// FB_TaktGenerator: 脉冲发生器
// 描述: 生成固定频率的方波脉冲信号 (50%占空比)

FUNCTION_BLOCK FB_TaktGenerator
VAR_INPUT
    Enable : BOOL;   // 使能信号 (TRUE=启用脉冲输出)
END_VAR
VAR_OUTPUT
    Takt_10Hz    : BOOL;  // 10Hz脉冲输出 (周期100ms)
    Takt_5Hz     : BOOL;  // 5Hz脉冲输出 (周期200ms)
    Takt_2_5Hz   : BOOL;  // 2.5Hz脉冲输出 (周期400ms)
    Takt_2Hz     : BOOL;  // 2Hz脉冲输出 (周期500ms)
    Takt_1_25Hz  : BOOL;  // 1.25Hz脉冲输出 (周期800ms)
    Takt_1Hz     : BOOL;  // 1Hz脉冲输出 (周期1s)
    Takt_0_625Hz : BOOL;  // 0.625Hz脉冲输出 (周期1.6s)
    Takt_0_5Hz   : BOOL;  // 0.5Hz脉冲输出 (周期2s)
    Takt_0_25Hz  : BOOL;  // 0.25Hz脉冲输出 (周期4s)
    Takt_0_2Hz   : BOOL;  // 0.2Hz脉冲输出 (周期5s)
END_VAR
VAR
    Cnt_10Hz     : DINT := 0;
    Cnt_5Hz      : DINT := 0;
    Cnt_2_5Hz    : DINT := 0;
    Cnt_2Hz      : DINT := 0;
    Cnt_1_25Hz   : DINT := 0;
    Cnt_1Hz      : DINT := 0;
    Cnt_0_625Hz  : DINT := 0;
    Cnt_0_5Hz    : DINT := 0;
    Cnt_0_25Hz   : DINT := 0;
    Cnt_0_2Hz    : DINT := 0;
END_VAR

BEGIN
    IF #Enable THEN
        // 10Hz: 周期100ms (假设10ms/扫描周期, 半周期=5)
        #Cnt_10Hz := #Cnt_10Hz + 1;
        IF #Cnt_10Hz >= 5 THEN
            #Takt_10Hz := NOT #Takt_10Hz;
            #Cnt_10Hz := 0;
        END_IF;

        // 5Hz: 周期200ms (半周期=10)
        #Cnt_5Hz := #Cnt_5Hz + 1;
        IF #Cnt_5Hz >= 10 THEN
            #Takt_5Hz := NOT #Takt_5Hz;
            #Cnt_5Hz := 0;
        END_IF;

        // 2.5Hz: 周期400ms (半周期=20)
        #Cnt_2_5Hz := #Cnt_2_5Hz + 1;
        IF #Cnt_2_5Hz >= 20 THEN
            #Takt_2_5Hz := NOT #Takt_2_5Hz;
            #Cnt_2_5Hz := 0;
        END_IF;

        // 2Hz: 周期500ms (半周期=25)
        #Cnt_2Hz := #Cnt_2Hz + 1;
        IF #Cnt_2Hz >= 25 THEN
            #Takt_2Hz := NOT #Takt_2Hz;
            #Cnt_2Hz := 0;
        END_IF;

        // 1.25Hz: 周期800ms (半周期=40)
        #Cnt_1_25Hz := #Cnt_1_25Hz + 1;
        IF #Cnt_1_25Hz >= 40 THEN
            #Takt_1_25Hz := NOT #Takt_1_25Hz;
            #Cnt_1_25Hz := 0;
        END_IF;

        // 1Hz: 周期1000ms (半周期=50)
        #Cnt_1Hz := #Cnt_1Hz + 1;
        IF #Cnt_1Hz >= 50 THEN
            #Takt_1Hz := NOT #Takt_1Hz;
            #Cnt_1Hz := 0;
        END_IF;

        // 0.625Hz: 周期1600ms (半周期=80)
        #Cnt_0_625Hz := #Cnt_0_625Hz + 1;
        IF #Cnt_0_625Hz >= 80 THEN
            #Takt_0_625Hz := NOT #Takt_0_625Hz;
            #Cnt_0_625Hz := 0;
        END_IF;

        // 0.5Hz: 周期2000ms (半周期=100)
        #Cnt_0_5Hz := #Cnt_0_5Hz + 1;
        IF #Cnt_0_5Hz >= 100 THEN
            #Takt_0_5Hz := NOT #Takt_0_5Hz;
            #Cnt_0_5Hz := 0;
        END_IF;

        // 0.25Hz: 周期4000ms (半周期=200)
        #Cnt_0_25Hz := #Cnt_0_25Hz + 1;
        IF #Cnt_0_25Hz >= 200 THEN
            #Takt_0_25Hz := NOT #Takt_0_25Hz;
            #Cnt_0_25Hz := 0;
        END_IF;

        // 0.2Hz: 周期5000ms (半周期=250)
        #Cnt_0_2Hz := #Cnt_0_2Hz + 1;
        IF #Cnt_0_2Hz >= 250 THEN
            #Takt_0_2Hz := NOT #Takt_0_2Hz;
            #Cnt_0_2Hz := 0;
        END_IF;
    ELSE
        // 禁用时复位所有输出和计数器
        #Takt_10Hz := FALSE;
        #Takt_5Hz := FALSE;
        #Takt_2_5Hz := FALSE;
        #Takt_2Hz := FALSE;
        #Takt_1_25Hz := FALSE;
        #Takt_1Hz := FALSE;
        #Takt_0_625Hz := FALSE;
        #Takt_0_5Hz := FALSE;
        #Takt_0_25Hz := FALSE;
        #Takt_0_2Hz := FALSE;
        #Cnt_10Hz := 0;
        #Cnt_5Hz := 0;
        #Cnt_2_5Hz := 0;
        #Cnt_2Hz := 0;
        #Cnt_1_25Hz := 0;
        #Cnt_1Hz := 0;
        #Cnt_0_625Hz := 0;
        #Cnt_0_5Hz := 0;
        #Cnt_0_25Hz := 0;
        #Cnt_0_2Hz := 0;
    END_IF;

END_FUNCTION_BLOCK
